(*
 * Simulacion_Trifasico_MPC_v8_M6_reducido_S71200.scl
 *
 * MPC REDUCIDO para S7-1200 (CPU 1212C). Base: Simulacion_Trifasico_MPC_v8_M6_it10_opt_S71200_v2.scl
 * (Parametros_MPC_v8: Ts = 0.1 s, P = 200, M = 6, mismos pesos y mismo filtro de Kalman).
 *
 * En la 1212C, el QP con restricciones (19 variables, 72 restricciones, solver KWIK) tardo de
 * 2 a mas de 12 s por ejecucion. Esta version conserva el estimador, el termino lineal del QP y
 * los limites del MPC, pero sustituye el QP por su solucion sin restricciones:
 *     zopt = -Hinv * f   (solo los movimientos u(k) de las 3 valvulas)
 * y despues recorta SIEMPRE con mpc_clipping (cambio por muestra 3.5 / 1.5 / 3 %, apertura 2-99 %).
 *  - Cuando ninguna restriccion esta activa, la accion es la misma que la del MPC completo
 *    (misma cuenta que la rama sin restricciones del QP).
 *  - Cuando hay restricciones activas (valvulas saturadas o limitadas en su cambio), el resultado
 *    puede diferir: el recorte no redistribuye la accion entre valvulas como el QP.
 * Sin QP ya no se usan qr, xgemv, xgerc, DropConstraint, abs_g, b_abs, maximum2, maximum, mtimes,
 * xnrm2, b_norm ni rt_floord: borrarlos del proyecto de TIA despues de importar.
 * LLAMAR DESDE UN OB CICLICO DE 100 ms. Requiere el DB global Diag_HIL.
 * [DIAG] Mediciones de RUNTIME <= 0.0 (vuelta del contador interno) se descartan.
 *)
DATA_BLOCK PLCGlobalVarMPC
STRUCT
    plc_ts_counter_MPC: DINT;
END_STRUCT
BEGIN
END_DATA_BLOCK
FUNCTION_BLOCK mpc_clipping_MPC
VAR_INPUT
    uk: ARRAY [0..2] OF REAL;
    uk1: ARRAY [0..2] OF REAL;
    b_uoff: ARRAY [0..2] OF REAL;
    b_ny: DINT;
    b_degrees: DINT;
END_VAR
VAR_OUTPUT
    uk_clipped: ARRAY [0..2] OF REAL;
END_VAR
VAR_IN_OUT
    b_Mlim: ARRAY [0..71] OF REAL;   (* solo lectura *)
    b_Mrows: ARRAY [0..71] OF DINT;  (* solo lectura *)
END_VAR
VAR
    nylim: DINT;
    umax: ARRAY [0..2] OF REAL;
    umin: ARRAY [0..2] OF REAL;
    dumin: ARRAY [0..2] OF REAL;
    dumax: ARRAY [0..2] OF REAL;
    iu: DINT;
    du: REAL;
    b_i: DINT;
    tmp: DINT;
    temp1: BOOL;
    temp2: BOOL;
    temp3: BOOL;
END_VAR
nylim := (400 * b_ny) + 1200;
uk_clipped[0] := uk[0];
umax[0] := 3.4028234663852886E+37;
umin[0] := -3.4028234663852886E+37;
dumin[0] := -3.4028234663852886E+37;
dumax[0] := 3.4028234663852886E+37;
uk_clipped[1] := uk[1];
umax[1] := 3.4028234663852886E+37;
umin[1] := -3.4028234663852886E+37;
dumin[1] := -3.4028234663852886E+37;
dumax[1] := 3.4028234663852886E+37;
uk_clipped[2] := uk[2];
umax[2] := 3.4028234663852886E+37;
umin[2] := -3.4028234663852886E+37;
dumin[2] := -3.4028234663852886E+37;
dumax[2] := 3.4028234663852886E+37;
FOR b_i := 0 TO 71 DO
    iu := b_Mrows[b_i];
    temp1 := FALSE;
    temp2 := FALSE;
    temp3 := FALSE;
    IF iu > (nylim - 1200) THEN
        IF iu <= (nylim - 1197) THEN
            iu := (iu - nylim) + 1199;
            umax[iu] := b_Mlim[b_i] + b_uoff[iu];
        ELSE
            temp3 := TRUE;
        END_IF;
    ELSE
        temp3 := TRUE;
    END_IF;
    IF temp3 THEN
        IF iu > (nylim - 600) THEN
            IF iu <= (nylim - 597) THEN
                iu := (iu - nylim) + 599;
                umin[iu] := ( -b_Mlim[b_i]) + b_uoff[iu];
            ELSE
                temp2 := TRUE;
            END_IF;
        ELSE
            temp2 := TRUE;
        END_IF;
    END_IF;
    IF temp2 THEN
        IF iu > nylim THEN
            IF iu <= (nylim + 3) THEN
                dumax[(iu - nylim) - 1] := b_Mlim[b_i];
            ELSE
                temp1 := TRUE;
            END_IF;
        ELSE
            temp1 := TRUE;
        END_IF;
    END_IF;
    IF temp1 THEN
        tmp := nylim + b_degrees;
        IF iu > (tmp - 1) THEN
            IF iu <= (tmp + 2) THEN
                dumin[(iu - nylim) - b_degrees] :=  -b_Mlim[b_i];
            END_IF;
        END_IF;
    END_IF;
END_FOR;
du := uk[0] - uk1[0];
IF du > dumax[0] THEN
    uk_clipped[0] := uk1[0] + dumax[0];
ELSIF du < dumin[0] THEN
    uk_clipped[0] := uk1[0] + dumin[0];
END_IF;
IF uk_clipped[0] > umax[0] THEN
    uk_clipped[0] := umax[0];
ELSIF uk_clipped[0] < umin[0] THEN
    uk_clipped[0] := umin[0];
END_IF;
du := uk[1] - uk1[1];
IF du > dumax[1] THEN
    uk_clipped[1] := uk1[1] + dumax[1];
ELSIF du < dumin[1] THEN
    uk_clipped[1] := uk1[1] + dumin[1];
END_IF;
IF uk_clipped[1] > umax[1] THEN
    uk_clipped[1] := umax[1];
ELSIF uk_clipped[1] < umin[1] THEN
    uk_clipped[1] := umin[1];
END_IF;
du := uk[2] - uk1[2];
IF du > dumax[2] THEN
    uk_clipped[2] := uk1[2] + dumax[2];
ELSIF du < dumin[2] THEN
    uk_clipped[2] := uk1[2] + dumin[2];
END_IF;
IF uk_clipped[2] > umax[2] THEN
    uk_clipped[2] := umax[2];
ELSIF uk_clipped[2] < umin[2] THEN
    uk_clipped[2] := umin[2];
END_IF;
END_FUNCTION_BLOCK
FUNCTION_BLOCK mpcblock_refmd_MPC
VAR_INPUT
    b_ref: ARRAY [0..2] OF REAL;
    b_yoff: ARRAY [0..2] OF REAL;
    b_RYscale: ARRAY [0..2] OF REAL;
END_VAR
VAR_OUTPUT
    rseq: ARRAY [0..2] OF REAL;   (* antes 0..599: solo se usan rseq[0..2] *)
    v: REAL;
END_VAR
VAR
    b_i: DINT;
    ref_0: REAL;
    ref_1: REAL;
    ref_2: REAL;
    b_RYscale_0: REAL;
    b_RYscale_1: REAL;
    b_RYscale_2: REAL;
    b_yoff_0: REAL;
    b_yoff_1: REAL;
    b_yoff_2: REAL;
END_VAR
ref_0 := b_ref[0];
ref_1 := b_ref[1];
ref_2 := b_ref[2];
b_RYscale_0 := b_RYscale[0];
b_RYscale_1 := b_RYscale[1];
b_RYscale_2 := b_RYscale[2];
b_yoff_0 := b_yoff[0];
b_yoff_1 := b_yoff[1];
b_yoff_2 := b_yoff[2];
FOR b_i := 0 TO 0 DO    (* solo rseq[0..2] se usa *)
    rseq[b_i * 3] := (ref_0 * b_RYscale_0) - b_yoff_0;
    rseq[(b_i * 3) + 1] := (ref_1 * b_RYscale_1) - b_yoff_1;
    rseq[(b_i * 3) + 2] := (ref_2 * b_RYscale_2) - b_yoff_2;
END_FOR;
v := 1.0;
END_FUNCTION_BLOCK
FUNCTION_BLOCK MPC_Control
VAR_INPUT
    ssMethodType: INT;
    moorx: ARRAY [0..2] OF REAL;
    b_ref: ARRAY [0..2] OF REAL;
END_VAR
VAR_OUTPUT
    mv: ARRAY [0..2] OF REAL;
END_VAR
VAR
    last_x_PreviousInput: ARRAY [0..6] OF REAL;
    last_mv_DSTATE: ARRAY [0..2] OF REAL;
    c_last_x_InitialCond: ARRAY [0..6] OF REAL := [0.47374550049727165,0.8,0.72,255106.009,0.0,0.0,0.0];
    MPC_3_b_myoff: ARRAY [0..2] OF REAL := [0.8,0.72,3.7];
    MPC_3_b_RYscale: ARRAY [0..2] OF REAL := [1.0,1.0,0.1];
    MPC_3_b_xoff: ARRAY [0..6] OF REAL := [0.47374550049727165,0.8,0.72,255106.009,0.0,0.0,0.0];
    b_a: ARRAY [0..20] OF REAL := [0.0,0.0,0.0,1.0,0.0,0.0,0.0,1.0,0.0,0.0,0.0,1.4503774389728313E-5,0.0,0.0,0.0,0.0,0.0,0.0,0.0,
        0.0,0.0];
    MPC_3_c_a: ARRAY [0..20] OF REAL := [-0.0772292027423523,0.12077646327456022,0.0038948707411090538,1352.9330397447068,
        3.4881337436777948,-1.3447885799979777,-1.1731438171327024,0.269035613232814,0.0038948707411099914,0.09786695730401461,
        348.05070726193321,0.11111867957141662,2.7949959088743932,-2.8155753844244291,0.059593437249509731,0.01962263557286395,
        0.0050480489343075492,14331.413461436903,1.6106730948140586,2.3311020292522353,2.408935193579286];
    MPC_3_b_Mlim: ARRAY [0..71] OF REAL := [0.333871875208127,0.752014397384409,0.515635973890735,0.333871875208127,
        0.752014397384409,0.515635973890735,0.333871875208127,0.752014397384409,0.515635973890735,0.333871875208127,0.752014397384409,
        0.515635973890735,0.333871875208127,0.752014397384409,0.515635973890735,0.333871875208127,0.752014397384409,0.515635973890735,
        0.636128124791873,0.21798560261559102,0.45436402610926496,0.636128124791873,0.21798560261559102,0.45436402610926496,
        0.636128124791873,0.21798560261559102,0.45436402610926496,0.636128124791873,0.21798560261559102,0.45436402610926496,
        0.636128124791873,0.21798560261559102,0.45436402610926496,0.636128124791873,0.21798560261559102,0.45436402610926496,0.035,0.015,
        0.03,0.035,0.015,0.03,0.035,0.015,0.03,0.035,0.015,0.03,0.035,0.015,0.03,0.035,0.015,0.03,0.035,0.015,0.03,0.035,0.015,
        0.03,0.035,0.015,0.03,0.035,0.015,0.03,0.035,0.015,0.03,0.035,0.015,0.03];
    MPC_3_b_Kx: ARRAY [0..125] OF REAL := [-7716.2321024491939,-10901.008671532656,-4264.9443651421188,0.001588040838629834,
        -2543.7442519006345,-1928.3474040587275,19.549174933816971,-44534.108859815329,-44494.776516572136,-26655.405567238093,
        0.0095121063518449449,-8398.6455416316712,-10368.267059564856,158.86185382546796,877.70571831208667,990.07022975809957,
        474.28108255756024,-0.0035701887162486057,96.5496604150103,99.981804413078876,-126.88330315000997,-7621.9188571763643,
        -10775.120625744157,-4206.5654308225376,0.0015700336455973293,-2519.1535379237243,-1907.0052261791157,19.280661326360363,
        -44188.119848216615,-44149.311125111242,-26390.969999054745,0.0094459267062587185,-8342.2703225681144,-10298.597291206755,
        157.85188650166057,864.95022738088733,975.66168439016542,466.81791298662728,-0.0035336819710021609,94.4868041100247,
        97.85316386731445,-125.93879584019494,-7528.1481322542822,-10649.931335099882,-4148.6767278274638,0.0015521046865827432,
        -2494.6400124657093,-1885.7587961853874,19.013959064141872,-43842.116288935795,-43803.826542255309,-26127.843886728973,
        0.0093796925467878947,-8285.8873550992248,-10228.919297363989,156.8419334382582,852.3095979437818,961.384106890396,459.43616436780036,
        -0.003497369852713806,92.447632839384539,95.74911914998566,-124.99418234183436,-7434.9230075303494,-10525.443894660129,
        -4091.2769580451954,0.0015342547665065048,-2470.2045128943837,-1864.6086925692725,18.749068146716176,-43496.122480806749,
        -43458.347088410825,-25866.027371158609,0.0093134067140901722,-8229.4967444644935,-10159.23320514503,155.83198146211291,
        839.78359704931961,947.23718912342133,452.13534732790527,-0.0034612522993006938,90.432068275420264,93.669582511506164,
        -124.04951211934259,-7342.2465048437853,-10401.661341488485,-4034.3648155478659,0.0015164846849855819,-2445.8478788030538,
        -1843.5554965261258,18.485988665509439,-43150.162591337648,-43112.896952629555,-25605.520593125708,0.0092470720701684772,
        -8173.0986508239621,-10089.539209226115,154.82201815145478,827.37198501561852,933.22061617028339,444.91497290855955,
        -0.0034253292477243787,88.440031602080353,91.614465843510473,-123.10483463065196,-7250.1215881048793,-10278.586654731167,
        -3977.9389865477651,0.00149879523623798,-2421.5709518529893,-1822.5997917608677,18.224720801734843,-42804.2606574284,
        -42767.500193326021,-25346.323693295184,0.0091806914982297729,-8116.6932889508143,-10019.83757147498,153.81203184149854,
        815.07451548496078,919.33406638300414,437.7745525706747,-0.0033896006339887937,86.47144350229388,89.5836806634611,
        -122.16019932703135];
    MPC_3_b_Ku1: ARRAY [0..53] OF REAL := [532.9519035819452,1758.7630386838541,-20.218495148255496,1758.7630386838541,
        9920.4082612993716,-164.30092992093171,-20.218495148255496,-164.30092992093171,131.49311423922407,527.80102628666316,
        1737.934860701725,-19.940788232849528,1746.9574860985949,9846.5918503106168,-163.25638356511735,-19.786511752201875,
        -161.71101778484783,130.514941055735,522.666313063715,1717.21838942958,-19.664954679108821,1735.1503109173054,9772.77075083077,
        -162.21185195795246,-19.359488246736596,-159.14605147852319,129.53665804804106,517.54793926655793,1696.6142696551719,
        -19.390994486572826,1723.3415351782228,9698.9487212665517,-161.16732147527,-18.93740822923742,-156.60596908182839,128.55831637410802,
        512.44608071469349,1676.1231380934234,-19.118907749797927,1711.5311924205112,9625.129520129678,-160.12277927000616,
        -18.520255194809877,-154.09070753671722,127.57996718519767,507.36091366067569,1655.7456233405144,-18.848694656201634,
        1699.7193276198914,9551.3169060341625,-159.07821327799945,-18.108012533640888,-151.60020265098143,126.60166162568011];
    MPC_3_b_Kr: ARRAY [0..53] OF REAL := [3186.8373350513389,4275.3677914960599,51.13509990647421,-32.452540397628589,26714.198696645544,72.918687149547608,
        -112.44555961175674,-475.25673471668864,252.72878690712173,3155.2425613858004,4216.8654170260106,50.638144210838703,
        -31.975100691061328,26449.325655557303,72.210143687081711,-110.79080635121332,-467.77820186026861,250.27164490947899,
        3123.8040857581582,4158.8539359264387,50.143499486122451,-31.502311016836352,26185.762042540995,71.504893608304656,
        -109.15217877028672,-460.38123779321489,247.82594499281888,3092.5219240585361,4101.3320539069082,49.651167400702548,
        -31.034149716397167,25923.508020768073,70.802939302930895,-107.52960162200367,-453.06535277614643,245.39169524300604,
        3061.396092190324,4044.2984688129827,49.161149624113243,-30.57059511536292,25662.563753294817,70.104283162373875,
        -105.92299960583885,-445.83005747772961,242.96890375165114,3030.4266060701984,3987.7518705822636,48.673447827046601,
        -30.111625523516803,25402.929403061011,69.408927579747242,-104.33229736767574,-438.67486297920362,240.55757861611488];   (* Kr reducida 18x3 *)
    (* Hinv3[3*j + c] = Hinv[19*j + c]: columnas de Hinv para los movimientos u(k) de las 3 valvulas *)
    MPC_3_b_Hinv3: ARRAY [0..56] OF REAL := [0.1702344980572631,-0.000316051953237396,-0.0001214533827540456,-0.000316051953237396,0.010547207252793461,
        2.1132487152157335E-5,-0.0001214533827540456,2.1132487152157335E-5,0.30304411821884769,-0.036345548841276047,
        -0.0001808791608454948,-6.514990994147179E-5,-0.00022994447282000675,-0.0023314158969080174,2.1728353827661485E-5,
        -7.8535204077971989E-5,1.0330320315621911E-5,-0.064405415788092474,-0.035434727013087031,-4.9534035220164727E-5,
        -8.97885060327611E-6,-0.00014382977097906262,-0.0022413766833578007,2.2273463510311548E-5,-3.4945956300716842E-5,
        1.2191170747377299E-7,-0.062989706993492336,-0.034542309014010772,7.8036147649309862E-5,4.65603793551569E-5,
        -5.7720706811642746E-5,-0.0021522792952646508,2.2723267969727878E-5,8.813456011776322E-6,-9.54953740575078E-6,
        -0.061614542822731315,-0.03366968301464044,0.00020190252942289518,0.00010110834451599296,2.8361008307101794E-5,
        -0.0020644122541486152,2.3046591530932414E-5,5.2380161360600679E-5,-1.8729858790232883E-5,-0.060282635561179215,
        -0.032817675154182616,0.0003221473455128597,0.00015444098334013595,0.00011438593593406882,-0.0019779594821308214,
        2.322473034505095E-5,9.552481608298865E-5,-2.7454115420488076E-5,-0.058995530723217567,0.0,0.0,0.0];
    MPC_3_b_uoff: ARRAY [0..2] OF REAL := [0.656128124791873,0.237985602615591,0.474364026109265];
    MPC_3_b_Mrows: ARRAY [0..71] OF DINT := [1201,1202,1203,1204,1205,1206,1207,1208,1209,1210,1211,1212,1213,1214,1215,1216,1217,
        1218,1801,1802,1803,1804,1805,1806,1807,1808,1809,1810,1811,1812,1813,1814,1815,1816,1817,1818,2401,2402,2403,2404,
        2405,2406,2407,2408,2409,2410,2411,2412,2413,2414,2415,2416,2417,2418,2419,2420,2421,2422,2423,2424,2425,2426,2427,
        2428,2429,2430,2431,2432,2433,2434,2435,2436];
    MPC_3_f_a: ARRAY [0..20] OF REAL := [1.322628327144006E-6,-0.00048116811531683895,-4.3296165052708516E-6,-55.375904267141834,
        0.0,0.0,0.0,-6.9150559684644062E-11,3.7716284508284807E-8,-0.0027971712823564414,-78.996564422017926,0.0,0.0,0.0,
        -2.394037186466665E-10,1.3057639972340998E-7,2.8628831792336135E-7,-273.49234867499621,0.0,0.0,0.0];
    MPC_3_g_a: ARRAY [0..20] OF REAL := [-0.0812759988320282,0.12878974211545094,0.004723574350295019,1608.467976495617,
        3.4881337436777868,-1.3447885799979735,-1.1731438171326984,0.27540380820784305,0.004147779263663315,0.10291146104511424,
        371.46041919189759,0.11111867957141465,2.7949959088743945,-2.8155753844244238,0.065710282048828311,0.023308594370287667,
        0.00655318586773693,16000.578760709672,1.6106730948139927,2.3311020292522739,2.4089351935793255];
    MPC_3_e_a: ARRAY [0..48] OF REAL := [0.9945076508163887,-7.4955911032675407E-6,0.018219343923005435,-0.86686845021470726,0.0,
        0.0,0.0,-0.0054923962532121753,0.99999067551082088,0.018219326989996565,-1.077349693812959,0.0,0.0,0.0,
        -4.0627503649808205E-13,2.2159162199695515E-10,0.99998342284905262,-0.4641225044555104,0.0,0.0,0.0,2.6237854624951297E-12,
        -9.54430195553142E-10,-2.0954813586927272E-9,0.99929334159686478,0.0,0.0,0.0,-6.3159654022047717E-6,0.0022977287773259252,
        2.0675277771461239E-5,264.43732399282771,1.0,0.0,0.0,0.002815004563879495,-1.3684281447907272E-7,2.54613431540441E-5,264.43733847702208,
        0.0,1.0,0.0,2.3147841327022809E-10,-1.26253752403586E-7,-2.7681092818992033E-7,264.43856123334115,0.0,0.0,1.0];
    i0_mpcblock_refmd: mpcblock_refmd_MPC;
    i0_mpc_clipping: mpc_clipping_MPC;
    xk: ARRAY [0..6] OF REAL;
    y_innov: ARRAY [0..2] OF REAL;
    v: REAL;
    rseq: ARRAY [0..2] OF REAL;
    zopt: ARRAY [0..2] OF REAL;
    b_i: DINT;
    rMin: REAL;
    tmp: DINT;
    kDrop: DINT;
    Xnorm0: REAL;
    cMin: REAL;
    cVal: REAL;
    z: ARRAY [0..18] OF REAL;
    t: REAL;
    j_k: DINT;
    rtb_xest: ARRAY [0..6] OF REAL;
    old_u: ARRAY [0..2] OF REAL;
    y_innov_0: REAL;
    D_tmp: DINT;
END_VAR
CASE ssMethodType OF
    0:
        PLCGlobalVarMPC.plc_ts_counter_MPC := 0;
        last_mv_DSTATE[0] := 0.656128124791873;
        last_mv_DSTATE[1] := 0.23798560261559079;
        last_mv_DSTATE[2] := 0.47436402610926476;
        FOR kDrop := 0 TO 6 DO
            last_x_PreviousInput[kDrop] := c_last_x_InitialCond[kDrop];
        END_FOR;
    1:
        IF PLCGlobalVarMPC.plc_ts_counter_MPC = 0 THEN
            (* [DIAG] inicio de la medicion *)
            "Diag_HIL".mpc_aux := RUNTIME("Diag_HIL".mpc_mem);

            (* Referencias escaladas *)
            i0_mpcblock_refmd(b_ref := b_ref, b_yoff := MPC_3_b_myoff, b_RYscale := MPC_3_b_RYscale);
            rseq := i0_mpcblock_refmd.rseq;
            v := i0_mpcblock_refmd.v;
            rMin := last_mv_DSTATE[0] - 0.656128124791873;
            Xnorm0 := last_mv_DSTATE[1] - 0.237985602615591;
            cMin := last_mv_DSTATE[2] - 0.474364026109265;

            (* Estimador: innovacion y estado corregido (sin cambios) *)
            FOR kDrop := 0 TO 6 DO
                xk[kDrop] := last_x_PreviousInput[kDrop] - MPC_3_b_xoff[kDrop];
            END_FOR;
            FOR j_k := 0 TO 2 DO
                cVal := 0.0;
                FOR D_tmp := 0 TO 6 DO
                    cVal := (b_a[(3 * D_tmp) + j_k] * xk[D_tmp]) + cVal;
                END_FOR;
                y_innov[j_k] := ((moorx[j_k] * MPC_3_b_RYscale[j_k]) - MPC_3_b_myoff[j_k]) - cVal;
            END_FOR;
            cVal := y_innov[1];
            t := y_innov[0];
            y_innov_0 := y_innov[2];
            FOR j_k := 0 TO 6 DO
                rtb_xest[j_k] := (((MPC_3_c_a[j_k + 7] * cVal) + (MPC_3_c_a[j_k] * t)) + (MPC_3_c_a[j_k + 14] * y_innov_0)
                    ) + xk[j_k];
            END_FOR;

            (* Termino lineal f del QP (z), igual que en el MPC completo *)
            FOR kDrop := 0 TO 18 DO
                z[kDrop] := 0.0;
            END_FOR;
            FOR b_i := 0 TO 17 DO
                cVal := 0.0;
                FOR j_k := 0 TO 6 DO
                    cVal := (MPC_3_b_Kx[(7 * b_i) + j_k] * rtb_xest[j_k]) + cVal;
                END_FOR;
                t := ((MPC_3_b_Kr[3 * b_i] * rseq[0]) + (MPC_3_b_Kr[(3 * b_i) + 1] * rseq[1])) + (MPC_3_b_Kr[(3 * b_i) + 2] * rseq[2]);
                z[b_i] := (((MPC_3_b_Ku1[(3 * b_i) + 1] * Xnorm0) + (MPC_3_b_Ku1[3 * b_i] * rMin)) + (MPC_3_b_Ku1[(3 * b_i)
                     + 2] * cMin)) + (cVal + t);
            END_FOR;

            (* MPC REDUCIDO: en lugar del QP con restricciones, la solucion sin restricciones
               zopt = -Hinv*f, solo para los movimientos u(k) de las 3 valvulas. Es la misma
               cuenta que hace el QP completo cuando ninguna restriccion esta activa. *)
            FOR tmp := 0 TO 2 DO
                Xnorm0 := 0.0;
                FOR j_k := 0 TO 18 DO
                    Xnorm0 := (( -MPC_3_b_Hinv3[(3 * j_k) + tmp]) * z[j_k]) + Xnorm0;
                END_FOR;
                zopt[tmp] := Xnorm0;
            END_FOR;
            b_i := 1;

            (* [DIAG] sin QP: estado 1, una "iteracion" *)
            "Diag_HIL".mpc_qp_estado := b_i;
            "Diag_HIL".mpc_iter_max := MAX(IN1 := "Diag_HIL".mpc_iter_max, IN2 := b_i);

            mv[0] := ((last_mv_DSTATE[0] - 0.656128124791873) + zopt[0]) + 0.656128124791873;
            mv[1] := ((last_mv_DSTATE[1] - 0.237985602615591) + zopt[1]) + 0.237985602615591;
            mv[2] := ((last_mv_DSTATE[2] - 0.474364026109265) + zopt[2]) + 0.474364026109265;
            (* Recorte SIEMPRE a los limites del MPC: cambio por muestra (3.5 / 1.5 / 3 %)
               y apertura (2-99 %), con el mismo bloque que usa el MPC completo *)
            old_u[0] := (last_mv_DSTATE[0] - 0.656128124791873) + 0.656128124791873;
            old_u[1] := (last_mv_DSTATE[1] - 0.237985602615591) + 0.237985602615591;
            old_u[2] := (last_mv_DSTATE[2] - 0.474364026109265) + 0.474364026109265;
            i0_mpc_clipping(uk := mv, uk1 := old_u, b_uoff := MPC_3_b_uoff, b_Mlim := MPC_3_b_Mlim, b_Mrows := MPC_3_b_Mrows,
                b_ny := 3, b_degrees := 19);
            mv := i0_mpc_clipping.uk_clipped;

            (* Actualizacion del estimador con la apertura aplicada (sin cambios) *)
            last_mv_DSTATE[0] := mv[0];
            rMin := mv[0] - 0.656128124791873;
            last_mv_DSTATE[1] := mv[1];
            Xnorm0 := mv[1] - 0.237985602615591;
            cMin := mv[2];
            last_mv_DSTATE[2] := mv[2];
            FOR j_k := 0 TO 6 DO
                cVal := 0.0;
                FOR D_tmp := 0 TO 6 DO
                    cVal := (MPC_3_e_a[(7 * D_tmp) + j_k] * xk[D_tmp]) + cVal;
                END_FOR;
                last_x_PreviousInput[j_k] := (((((MPC_3_f_a[j_k + 7] * Xnorm0) + (MPC_3_f_a[j_k] * rMin)) + (MPC_3_f_a[j_k + 14] * (cMin - 0.474364026109265)
                    )) + cVal) + (((MPC_3_g_a[j_k + 7] * y_innov[1]) + (MPC_3_g_a[j_k] * y_innov[0])) + (MPC_3_g_a[j_k + 14] * y_innov[2])
                    )) + MPC_3_b_xoff[j_k];
            END_FOR;

            (* [DIAG] fin de la medicion: tiempo de esta ejecucion en ms *)
            "Diag_HIL".mpc_ms := RUNTIME("Diag_HIL".mpc_mem) * 1000.0;

            (* [DIAG] reinicio de estadisticas desde la tabla de observacion *)
            IF "Diag_HIL".mpc_reset THEN
                "Diag_HIL".mpc_n := 0;
                "Diag_HIL".mpc_sum_ms := 0.0;
                "Diag_HIL".mpc_max_ms := 0.0;
                "Diag_HIL".mpc_iter_max := 0;
                "Diag_HIL".mpc_n_tope := 0;
                "Diag_HIL".mpc_n_infactible := 0;
                "Diag_HIL".mpc_reset := FALSE;
            END_IF;

            (* [DIAG] promedio y maximo desde el ultimo reset *)
            (* [DIAG] Si el contador interno de RUNTIME da la vuelta, la medicion sale <= 0.0 y
               Siemens indica descartarla: solo se acumulan mediciones positivas. *)
            IF "Diag_HIL".mpc_ms > 0.0 THEN
                "Diag_HIL".mpc_n := "Diag_HIL".mpc_n + 1;
                "Diag_HIL".mpc_sum_ms := "Diag_HIL".mpc_sum_ms + "Diag_HIL".mpc_ms;
                "Diag_HIL".mpc_prom_ms := "Diag_HIL".mpc_sum_ms / DINT_TO_LREAL("Diag_HIL".mpc_n);
                "Diag_HIL".mpc_max_ms := MAX(IN1 := "Diag_HIL".mpc_max_ms, IN2 := "Diag_HIL".mpc_ms);
            END_IF;
        END_IF;
        IF PLCGlobalVarMPC.plc_ts_counter_MPC >= 0 THEN   (* divisor desactivado: OB de 100 ms *)
            PLCGlobalVarMPC.plc_ts_counter_MPC := 0;
        ELSE
            PLCGlobalVarMPC.plc_ts_counter_MPC := PLCGlobalVarMPC.plc_ts_counter_MPC + 1;
        END_IF;
END_CASE;
END_FUNCTION_BLOCK
